Fanuc KAREL source: KO00005.KL

PROGRAM KO00005
%NOLOCKGROUP
VAR
  P1: POSITION
  P2: POSITION
  P3: POSITION
  P4: POSITION
  OUT: POSITION
BEGIN
  OUT = FRAME(P1, P2, P3, P4)
END KO00005
